TYPE "ST_PressDemoLineConfig"
VERSION : 0.1
   STRUCT
      "SchemaVersion" : UInt := 1;
      "UtcOffsetMin" : DInt;
      "ShiftStartMin" : Array[1..5] of DInt;
      "ShiftDurationMin" : Array[1..5] of DInt;
      "ShiftActiveDays" : Array[1..5] of DInt;
      "ShiftTarget" : Array[1..5] of DInt;
   END_STRUCT;
END_TYPE
